(* IEC 61131-3 sources: RAG_PLC/data/result/test/062, 2 files *)

(* ---- wrapped.st ---- *)
(* =========================================================
   Generated by PLC-Eval Benchmark Wrapper
   ========================================================= *)

FUNCTION_BLOCK LLM_Wrapper_FB
VAR_INPUT
    I0 : BOOL;
    I1 : BOOL;
    I2 : BOOL;
    I3 : BOOL;
    MAN : BOOL;
    STP : BOOL;
    M0 : BOOL;
    M1 : BOOL;
    M2 : BOOL;
    M3 : BOOL;
END_VAR

VAR_OUTPUT
    Q0 : BOOL;
    Q1 : BOOL;
    Q2 : BOOL;
    Q3 : BOOL;
    STATUS : BYTE;
END_VAR

VAR
    edge : BOOL;
    pos : INT;
    tog : BOOL;
END_VAR

(*@KEY@: WORKSHEET
NAME: MANUAL_4
IEC_LANGUAGE: ST
*)
IF man THEN
    IF NOT TOG THEN
        Q0 := M0;
        Q1 := M1;
        Q2 := M2;
        Q3 := M3;
        STATUS := BYTE#101;
    END_IF;
    IF STP AND NOT edge THEN
        tog := TRUE;
        CASE pos OF
            0: Q0 := TRUE;
                Q1 := FALSE;
                Q2 := FALSE;
                Q3 := FALSE;
                STATUS := BYTE#110;
            1: Q0 := FALSE;
                Q1 := TRUE;
                Q2 := FALSE;
                Q3 := FALSE;
                STATUS := BYTE#111;
            2: Q0 := FALSE;
                Q1 := FALSE;
                Q2 := TRUE;
                Q3 := FALSE;
                STATUS := BYTE#112;
            3: Q0 := FALSE;
                Q1 := FALSE;
                Q2 := FALSE;
                Q3 := TRUE;
                STATUS := BYTE#113;
        END_CASE;
        pos := INC(pos,1,3);
    END_IF;
ELSE
    Q0 := I0;
    Q1 := I1;
    Q2 := I2;
    Q3 := I3;
    STATUS := BYTE#100;
    tog := FALSE;
    pos := 0;
END_IF;

(* 记住 STP 信号的状态 *)
edge := STP;
END_FUNCTION_BLOCK

PROGRAM Auto_Proxy_Prg
  VAR
    instance : LLM_Wrapper_FB;
  END_VAR

  instance();
END_PROGRAM

CONFIGURATION Config0
  RESOURCE Res0 ON PLC
    TASK TaskMain(INTERVAL := T#20ms, PRIORITY := 0);
    PROGRAM Inst0 WITH TaskMain : Auto_Proxy_Prg;
  END_RESOURCE
END_CONFIGURATION

(* ---- raw_code.st ---- *)
VAR_INPUT
    I0 : BOOL;
    I1 : BOOL;
    I2 : BOOL;
    I3 : BOOL;
    MAN : BOOL;
    STP : BOOL;
    M0 : BOOL;
    M1 : BOOL;
    M2 : BOOL;
    M3 : BOOL;
END_VAR

VAR_OUTPUT
    Q0 : BOOL;
    Q1 : BOOL;
    Q2 : BOOL;
    Q3 : BOOL;
    STATUS : BYTE;
END_VAR

VAR
    edge : BOOL;
    pos : INT;
    tog : BOOL;
END_VAR

(*@KEY@: WORKSHEET
NAME: MANUAL_4
IEC_LANGUAGE: ST
*)
IF man THEN
    IF NOT TOG THEN
        Q0 := M0;
        Q1 := M1;
        Q2 := M2;
        Q3 := M3;
        STATUS := BYTE#101;
    END_IF;
    IF STP AND NOT edge THEN
        tog := TRUE;
        CASE pos OF
            0: Q0 := TRUE;
                Q1 := FALSE;
                Q2 := FALSE;
                Q3 := FALSE;
                STATUS := BYTE#110;
            1: Q0 := FALSE;
                Q1 := TRUE;
                Q2 := FALSE;
                Q3 := FALSE;
                STATUS := BYTE#111;
            2: Q0 := FALSE;
                Q1 := FALSE;
                Q2 := TRUE;
                Q3 := FALSE;
                STATUS := BYTE#112;
            3: Q0 := FALSE;
                Q1 := FALSE;
                Q2 := FALSE;
                Q3 := TRUE;
                STATUS := BYTE#113;
        END_CASE;
        pos := INC(pos,1,3);
    END_IF;
ELSE
    Q0 := I0;
    Q1 := I1;
    Q2 := I2;
    Q3 := I3;
    STATUS := BYTE#100;
    tog := FALSE;
    pos := 0;
END_IF;

(* 记住 STP 信号的状态 *)
edge := STP;
